(* IEC 61131-3 sources: plc-hackathon-2026/work/dump/MyController/Plc Logic/Application, 7 files *)

(* ---- SimCal.st ---- *)
// DATA_BLOCK "SimCal"
// NON_RETAIN
// Kumulativni dani po mjesecima (nepr. godina)
   VAR_GLOBAL
      CumDays : Array[0..12] of Int;
   END_VAR

(* ---- SimCtrl.st ---- *)
// DATA_BLOCK "SimCtrl"
// { S7_Optimized_Access := 'TRUE' }
// VERSION : 0.1
// NON_RETAIN
// ---------------------------------------------------------------------
// Upravljanje simulacijom (HMI/organizator)
// ---------------------------------------------------------------------
   VAR_GLOBAL
      run : Bool;   // TRUE = simulacija radi (pauza = FALSE)
      reset : Bool;   // 1 = reinicijalizacija (obradi se u OB30, sam se vraca na FALSE)
      price_mode : Int;   // 0 = dvotarifno, 1 = dan-unaprijed
      k : DInt;   // trenutni korak
      finished : BOOL;   // { ExternalWritable := 'False'}
      tripped : BOOL;   // { ExternalWritable := 'False'}
      stepActive : Bool;   // postavlja Sim_Core faza 1 --- promjena cycle timea (tvoja mreza SET_CINT) ---
      cycle_time_ms : UDInt;
      cycle_time_us : UDINT;   // { ExternalAccessible := 'False'; ExternalVisible := 'False'; ExternalWritable := 'False'}
      change_cycle : Bool;   // HMI: 1 -> primijeni cycle_time_ms
      change_cycle_P1 : BOOL;   // { ExternalAccessible := 'False'; ExternalVisible := 'False'; ExternalWritable := 'False'} memorijski bit za P_TRIG
      ret_val_cint : UDInt;   // { ExternalAccessible := 'False'; ExternalVisible := 'False'; ExternalWritable := 'False'}
   END_VAR

(* ---- SimIO.st ---- *)
// DATA_BLOCK "SimIO"
// { S7_Optimized_Access := 'TRUE' }
// VERSION : 0.1
// NON_RETAIN
// ---------------------------------------------------------------------
// Razmjena regulator <-> simulator
// ---------------------------------------------------------------------
   VAR_GLOBAL
      simOut : typeSimOut;
      simCmd : typeSimCmd;
   END_VAR

(* ---- SimParam.st ---- *)
// DATA_BLOCK "SimParam"
// NON_RETAIN
// ---------------------------------------------------------------------
// Globalni parametri
// ---------------------------------------------------------------------
   VAR_GLOBAL
      TS_H : Real;
      SIM_YEAR : UInt;   // neprijestupna godina (365 d = 35040 koraka)
      START_WEEKDAY : Int;   // 1.1.2025. = srijeda (1=pon)
      FNE_MAX_POWER : Real;
      BESS_CAPACITY : Real;
      BESS_MAX_CHG : Real;
      BESS_MAX_DCH : Real;
      BESS_SOC_MIN : Real;   // (*) sigurnosna donja granica [%]
      BESS_SOC_MAX : Real;   // (*) sigurnosna gornja granica [%]
      BESS_SOC_INIT : Real;   // (*)
      BESS_ETA_CHG : Real;   // (*)
      BESS_ETA_DCH : Real;   // (*)
      EV_MAX_CHARGE : Real;
      EV_ETA : Real;   // (*)
      EGC_MAX_IMPORT : Real;
      EGC_MAX_EXPORT : Real;   // --- tarife (*) - uskladi s HEP Bijeli / srednji napon --- cijena ENERGIJE dolazi iz profila (Prof_PriceTT / Prof_PriceDA, EUR/kWh); VT/NT iz Prof_VT
      GRID_VT : Real;   // mrezarina VT [EUR/kWh]  (HEP ODS, Bijeli 2, SN, od 1.1.2025.)
      GRID_NT : Real;   // mrezarina NT [EUR/kWh]
      PEAK_PRICE : Real;   // vrsna snaga [EUR/kW po mjesecu]
      EXPORT_FACTOR : Real;   // (*) izvoz se placa cijena_energije * faktor
   END_VAR

(* ---- SimScore.st ---- *)
// DATA_BLOCK "SimScore"
// NON_RETAIN
// Sluzbeni rezultat za ocjenjivanje (godisnji totali)
   VAR_GLOBAL
      total : typeAgg;
   END_VAR

(* ---- Team_Main.st ---- *)
FUNCTION_BLOCK Team_Main
VAR_INPUT
      simOut : typeSimOut;
END_VAR
VAR_OUTPUT
      simCmd : typeSimCmd;
END_VAR
VAR_TEMP

END_VAR

// ---IMPL---

(* ---- SR_Main_Sim.st ---- *)
PROGRAM SR_Main_Sim
VAR
	Init_Prof_EV_DB: Init_Prof_EV;
	Init_Prof_FEC_DB: Init_Prof_FEC;
	Init_Prof_FNE_DB: Init_Prof_FNE;
	Init_Prof_PriceDA_DB: Init_Prof_PriceDA;
	Init_Prof_PriceTT_DB: Init_Prof_PriceTT;
	Init_Prof_VT_DB: Init_Prof_VT;
	Init_SimCal_DB: Init_SimCal;
	Init_SimParam_DB: Init_SimParam;
	Init_SimCtrl_DB: Init_SimCtrl;
	Sim_Core_DB: Sim_Core;
	Team_Main_DB: Team_Main;
	Init_All_DB: Init_All;
	PLC_Started: BOOL;
	Datum_Vrijeme_Get_DB: Datum_Vrijeme_Get;
	Datum_Vrijeme_Set_DB: Datum_Vrijeme_Set;
END_VAR
